Fanuc KAREL source: KT00317.KL

PROGRAM KT00317
%NOLOCKGROUP
VAR
  P1: XYZWPR
  P2: XYZWPREXT
  OUT: BOOLEAN
BEGIN
  P1.X = 1.0
    P2.Y = 2.0
  OUT = P1 <> P2
END KT00317
